(* IEC 61131-3 sources: STAR-PLC-Agent/results/raw/four_group_20261114/star_terra/PUB011/generation/sim_00, 1 file *)

(* ---- test_program.st ---- *)
PROGRAM PLC_PRG
VAR
 BenchStep : UDINT := 0;
 BenchCalls : UDINT := 0;
 BenchDone : BOOL := FALSE;
 BenchUut0 : FB_Task;
 BenchUut1 : FB_Task;
 TraceIn_Mode : ARRAY[0..15] OF BOOL;
 TraceIn_ForwardButton : ARRAY[0..15] OF BOOL;
 TraceIn_ReverseButton : ARRAY[0..15] OF BOOL;
 TraceIn_SensorA : ARRAY[0..15] OF BOOL;
 TraceIn_SensorB : ARRAY[0..15] OF BOOL;
 TraceIn_SensorC : ARRAY[0..15] OF BOOL;
 TraceIn_ButtonA : ARRAY[0..15] OF BOOL;
 TraceIn_ButtonB : ARRAY[0..15] OF BOOL;
 TraceIn_ButtonC : ARRAY[0..15] OF BOOL;
 TraceOut_MotorForward : ARRAY[0..15] OF BOOL;
 TraceOut_MotorReverse : ARRAY[0..15] OF BOOL;
 TraceOut_CompletionLight : ARRAY[0..15] OF BOOL;
END_VAR

IF NOT BenchDone THEN
 CASE BenchStep OF
 0:
   BenchUut0.Mode := TRUE;
   BenchUut0.ForwardButton := FALSE;
   BenchUut0.ReverseButton := FALSE;
   BenchUut0.SensorA := TRUE;
   BenchUut0.SensorB := FALSE;
   BenchUut0.SensorC := FALSE;
   BenchUut0.ButtonA := FALSE;
   BenchUut0.ButtonB := FALSE;
   BenchUut0.ButtonC := FALSE;
   TraceIn_Mode[0] := BenchUut0.Mode;
   TraceIn_ForwardButton[0] := BenchUut0.ForwardButton;
   TraceIn_ReverseButton[0] := BenchUut0.ReverseButton;
   TraceIn_SensorA[0] := BenchUut0.SensorA;
   TraceIn_SensorB[0] := BenchUut0.SensorB;
   TraceIn_SensorC[0] := BenchUut0.SensorC;
   TraceIn_ButtonA[0] := BenchUut0.ButtonA;
   TraceIn_ButtonB[0] := BenchUut0.ButtonB;
   TraceIn_ButtonC[0] := BenchUut0.ButtonC;
   BenchUut0();
   TraceOut_MotorForward[0] := BenchUut0.MotorForward;
   TraceOut_MotorReverse[0] := BenchUut0.MotorReverse;
   TraceOut_CompletionLight[0] := BenchUut0.CompletionLight;
   BenchCalls := BenchCalls + 1;
 1:
   BenchUut0.Mode := TRUE;
   BenchUut0.ForwardButton := FALSE;
   BenchUut0.ReverseButton := FALSE;
   BenchUut0.SensorA := TRUE;
   BenchUut0.SensorB := FALSE;
   BenchUut0.SensorC := FALSE;
   BenchUut0.ButtonA := TRUE;
   BenchUut0.ButtonB := FALSE;
   BenchUut0.ButtonC := FALSE;
   TraceIn_Mode[1] := BenchUut0.Mode;
   TraceIn_ForwardButton[1] := BenchUut0.ForwardButton;
   TraceIn_ReverseButton[1] := BenchUut0.ReverseButton;
   TraceIn_SensorA[1] := BenchUut0.SensorA;
   TraceIn_SensorB[1] := BenchUut0.SensorB;
   TraceIn_SensorC[1] := BenchUut0.SensorC;
   TraceIn_ButtonA[1] := BenchUut0.ButtonA;
   TraceIn_ButtonB[1] := BenchUut0.ButtonB;
   TraceIn_ButtonC[1] := BenchUut0.ButtonC;
   BenchUut0();
   TraceOut_MotorForward[1] := BenchUut0.MotorForward;
   TraceOut_MotorReverse[1] := BenchUut0.MotorReverse;
   TraceOut_CompletionLight[1] := BenchUut0.CompletionLight;
   BenchCalls := BenchCalls + 1;
 2:
   BenchUut0.Mode := TRUE;
   BenchUut0.ForwardButton := FALSE;
   BenchUut0.ReverseButton := FALSE;
   BenchUut0.SensorA := FALSE;
   BenchUut0.SensorB := TRUE;
   BenchUut0.SensorC := FALSE;
   BenchUut0.ButtonA := FALSE;
   BenchUut0.ButtonB := TRUE;
   BenchUut0.ButtonC := FALSE;
   TraceIn_Mode[2] := BenchUut0.Mode;
   TraceIn_ForwardButton[2] := BenchUut0.ForwardButton;
   TraceIn_ReverseButton[2] := BenchUut0.ReverseButton;
   TraceIn_SensorA[2] := BenchUut0.SensorA;
   TraceIn_SensorB[2] := BenchUut0.SensorB;
   TraceIn_SensorC[2] := BenchUut0.SensorC;
   TraceIn_ButtonA[2] := BenchUut0.ButtonA;
   TraceIn_ButtonB[2] := BenchUut0.ButtonB;
   TraceIn_ButtonC[2] := BenchUut0.ButtonC;
   BenchUut0();
   TraceOut_MotorForward[2] := BenchUut0.MotorForward;
   TraceOut_MotorReverse[2] := BenchUut0.MotorReverse;
   TraceOut_CompletionLight[2] := BenchUut0.CompletionLight;
   BenchCalls := BenchCalls + 1;
 3:
   BenchUut0.Mode := TRUE;
   BenchUut0.ForwardButton := FALSE;
   BenchUut0.ReverseButton := FALSE;
   BenchUut0.SensorA := FALSE;
   BenchUut0.SensorB := TRUE;
   BenchUut0.SensorC := FALSE;
   BenchUut0.ButtonA := FALSE;
   BenchUut0.ButtonB := TRUE;
   BenchUut0.ButtonC := FALSE;
   TraceIn_Mode[3] := BenchUut0.Mode;
   TraceIn_ForwardButton[3] := BenchUut0.ForwardButton;
   TraceIn_ReverseButton[3] := BenchUut0.ReverseButton;
   TraceIn_SensorA[3] := BenchUut0.SensorA;
   TraceIn_SensorB[3] := BenchUut0.SensorB;
   TraceIn_SensorC[3] := BenchUut0.SensorC;
   TraceIn_ButtonA[3] := BenchUut0.ButtonA;
   TraceIn_ButtonB[3] := BenchUut0.ButtonB;
   TraceIn_ButtonC[3] := BenchUut0.ButtonC;
   BenchUut0();
   TraceOut_MotorForward[3] := BenchUut0.MotorForward;
   TraceOut_MotorReverse[3] := BenchUut0.MotorReverse;
   TraceOut_CompletionLight[3] := BenchUut0.CompletionLight;
   BenchCalls := BenchCalls + 1;
 4:
   BenchUut0.Mode := TRUE;
   BenchUut0.ForwardButton := FALSE;
   BenchUut0.ReverseButton := FALSE;
   BenchUut0.SensorA := FALSE;
   BenchUut0.SensorB := FALSE;
   BenchUut0.SensorC := TRUE;
   BenchUut0.ButtonA := FALSE;
   BenchUut0.ButtonB := FALSE;
   BenchUut0.ButtonC := TRUE;
   TraceIn_Mode[4] := BenchUut0.Mode;
   TraceIn_ForwardButton[4] := BenchUut0.ForwardButton;
   TraceIn_ReverseButton[4] := BenchUut0.ReverseButton;
   TraceIn_SensorA[4] := BenchUut0.SensorA;
   TraceIn_SensorB[4] := BenchUut0.SensorB;
   TraceIn_SensorC[4] := BenchUut0.SensorC;
   TraceIn_ButtonA[4] := BenchUut0.ButtonA;
   TraceIn_ButtonB[4] := BenchUut0.ButtonB;
   TraceIn_ButtonC[4] := BenchUut0.ButtonC;
   BenchUut0();
   TraceOut_MotorForward[4] := BenchUut0.MotorForward;
   TraceOut_MotorReverse[4] := BenchUut0.MotorReverse;
   TraceOut_CompletionLight[4] := BenchUut0.CompletionLight;
   BenchCalls := BenchCalls + 1;
 5:
   BenchUut0.Mode := TRUE;
   BenchUut0.ForwardButton := FALSE;
   BenchUut0.ReverseButton := FALSE;
   BenchUut0.SensorA := FALSE;
   BenchUut0.SensorB := FALSE;
   BenchUut0.SensorC := TRUE;
   BenchUut0.ButtonA := FALSE;
   BenchUut0.ButtonB := FALSE;
   BenchUut0.ButtonC := TRUE;
   TraceIn_Mode[5] := BenchUut0.Mode;
   TraceIn_ForwardButton[5] := BenchUut0.ForwardButton;
   TraceIn_ReverseButton[5] := BenchUut0.ReverseButton;
   TraceIn_SensorA[5] := BenchUut0.SensorA;
   TraceIn_SensorB[5] := BenchUut0.SensorB;
   TraceIn_SensorC[5] := BenchUut0.SensorC;
   TraceIn_ButtonA[5] := BenchUut0.ButtonA;
   TraceIn_ButtonB[5] := BenchUut0.ButtonB;
   TraceIn_ButtonC[5] := BenchUut0.ButtonC;
   BenchUut0();
   TraceOut_MotorForward[5] := BenchUut0.MotorForward;
   TraceOut_MotorReverse[5] := BenchUut0.MotorReverse;
   TraceOut_CompletionLight[5] := BenchUut0.CompletionLight;
   BenchCalls := BenchCalls + 1;
 6:
   BenchUut0.Mode := TRUE;
   BenchUut0.ForwardButton := FALSE;
   BenchUut0.ReverseButton := FALSE;
   BenchUut0.SensorA := FALSE;
   BenchUut0.SensorB := FALSE;
   BenchUut0.SensorC := TRUE;
   BenchUut0.ButtonA := FALSE;
   BenchUut0.ButtonB := FALSE;
   BenchUut0.ButtonC := FALSE;
   TraceIn_Mode[6] := BenchUut0.Mode;
   TraceIn_ForwardButton[6] := BenchUut0.ForwardButton;
   TraceIn_ReverseButton[6] := BenchUut0.ReverseButton;
   TraceIn_SensorA[6] := BenchUut0.SensorA;
   TraceIn_SensorB[6] := BenchUut0.SensorB;
   TraceIn_SensorC[6] := BenchUut0.SensorC;
   TraceIn_ButtonA[6] := BenchUut0.ButtonA;
   TraceIn_ButtonB[6] := BenchUut0.ButtonB;
   TraceIn_ButtonC[6] := BenchUut0.ButtonC;
   BenchUut0();
   TraceOut_MotorForward[6] := BenchUut0.MotorForward;
   TraceOut_MotorReverse[6] := BenchUut0.MotorReverse;
   TraceOut_CompletionLight[6] := BenchUut0.CompletionLight;
   BenchCalls := BenchCalls + 1;
 7:
   BenchUut0.Mode := TRUE;
   BenchUut0.ForwardButton := FALSE;
   BenchUut0.ReverseButton := FALSE;
   BenchUut0.SensorA := FALSE;
   BenchUut0.SensorB := FALSE;
   BenchUut0.SensorC := FALSE;
   BenchUut0.ButtonA := FALSE;
   BenchUut0.ButtonB := FALSE;
   BenchUut0.ButtonC := FALSE;
   TraceIn_Mode[7] := BenchUut0.Mode;
   TraceIn_ForwardButton[7] := BenchUut0.ForwardButton;
   TraceIn_ReverseButton[7] := BenchUut0.ReverseButton;
   TraceIn_SensorA[7] := BenchUut0.SensorA;
   TraceIn_SensorB[7] := BenchUut0.SensorB;
   TraceIn_SensorC[7] := BenchUut0.SensorC;
   TraceIn_ButtonA[7] := BenchUut0.ButtonA;
   TraceIn_ButtonB[7] := BenchUut0.ButtonB;
   TraceIn_ButtonC[7] := BenchUut0.ButtonC;
   BenchUut0();
   TraceOut_MotorForward[7] := BenchUut0.MotorForward;
   TraceOut_MotorReverse[7] := BenchUut0.MotorReverse;
   TraceOut_CompletionLight[7] := BenchUut0.CompletionLight;
   BenchCalls := BenchCalls + 1;
 8:
   BenchUut1.Mode := FALSE;
   BenchUut1.ForwardButton := TRUE;
   BenchUut1.ReverseButton := FALSE;
   BenchUut1.SensorA := FALSE;
   BenchUut1.SensorB := FALSE;
   BenchUut1.SensorC := FALSE;
   BenchUut1.ButtonA := FALSE;
   BenchUut1.ButtonB := FALSE;
   BenchUut1.ButtonC := FALSE;
   TraceIn_Mode[8] := BenchUut1.Mode;
   TraceIn_ForwardButton[8] := BenchUut1.ForwardButton;
   TraceIn_ReverseButton[8] := BenchUut1.ReverseButton;
   TraceIn_SensorA[8] := BenchUut1.SensorA;
   TraceIn_SensorB[8] := BenchUut1.SensorB;
   TraceIn_SensorC[8] := BenchUut1.SensorC;
   TraceIn_ButtonA[8] := BenchUut1.ButtonA;
   TraceIn_ButtonB[8] := BenchUut1.ButtonB;
   TraceIn_ButtonC[8] := BenchUut1.ButtonC;
   BenchUut1();
   TraceOut_MotorForward[8] := BenchUut1.MotorForward;
   TraceOut_MotorReverse[8] := BenchUut1.MotorReverse;
   TraceOut_CompletionLight[8] := BenchUut1.CompletionLight;
   BenchCalls := BenchCalls + 1;
 9:
   BenchUut1.Mode := FALSE;
   BenchUut1.ForwardButton := TRUE;
   BenchUut1.ReverseButton := TRUE;
   BenchUut1.SensorA := FALSE;
   BenchUut1.SensorB := FALSE;
   BenchUut1.SensorC := FALSE;
   BenchUut1.ButtonA := FALSE;
   BenchUut1.ButtonB := FALSE;
   BenchUut1.ButtonC := FALSE;
   TraceIn_Mode[9] := BenchUut1.Mode;
   TraceIn_ForwardButton[9] := BenchUut1.ForwardButton;
   TraceIn_ReverseButton[9] := BenchUut1.ReverseButton;
   TraceIn_SensorA[9] := BenchUut1.SensorA;
   TraceIn_SensorB[9] := BenchUut1.SensorB;
   TraceIn_SensorC[9] := BenchUut1.SensorC;
   TraceIn_ButtonA[9] := BenchUut1.ButtonA;
   TraceIn_ButtonB[9] := BenchUut1.ButtonB;
   TraceIn_ButtonC[9] := BenchUut1.ButtonC;
   BenchUut1();
   TraceOut_MotorForward[9] := BenchUut1.MotorForward;
   TraceOut_MotorReverse[9] := BenchUut1.MotorReverse;
   TraceOut_CompletionLight[9] := BenchUut1.CompletionLight;
   BenchCalls := BenchCalls + 1;
 10:
   BenchUut1.Mode := FALSE;
   BenchUut1.ForwardButton := FALSE;
   BenchUut1.ReverseButton := TRUE;
   BenchUut1.SensorA := FALSE;
   BenchUut1.SensorB := FALSE;
   BenchUut1.SensorC := FALSE;
   BenchUut1.ButtonA := FALSE;
   BenchUut1.ButtonB := FALSE;
   BenchUut1.ButtonC := FALSE;
   TraceIn_Mode[10] := BenchUut1.Mode;
   TraceIn_ForwardButton[10] := BenchUut1.ForwardButton;
   TraceIn_ReverseButton[10] := BenchUut1.ReverseButton;
   TraceIn_SensorA[10] := BenchUut1.SensorA;
   TraceIn_SensorB[10] := BenchUut1.SensorB;
   TraceIn_SensorC[10] := BenchUut1.SensorC;
   TraceIn_ButtonA[10] := BenchUut1.ButtonA;
   TraceIn_ButtonB[10] := BenchUut1.ButtonB;
   TraceIn_ButtonC[10] := BenchUut1.ButtonC;
   BenchUut1();
   TraceOut_MotorForward[10] := BenchUut1.MotorForward;
   TraceOut_MotorReverse[10] := BenchUut1.MotorReverse;
   TraceOut_CompletionLight[10] := BenchUut1.CompletionLight;
   BenchCalls := BenchCalls + 1;
 11:
   BenchUut1.Mode := TRUE;
   BenchUut1.ForwardButton := FALSE;
   BenchUut1.ReverseButton := TRUE;
   BenchUut1.SensorA := TRUE;
   BenchUut1.SensorB := FALSE;
   BenchUut1.SensorC := FALSE;
   BenchUut1.ButtonA := TRUE;
   BenchUut1.ButtonB := FALSE;
   BenchUut1.ButtonC := FALSE;
   TraceIn_Mode[11] := BenchUut1.Mode;
   TraceIn_ForwardButton[11] := BenchUut1.ForwardButton;
   TraceIn_ReverseButton[11] := BenchUut1.ReverseButton;
   TraceIn_SensorA[11] := BenchUut1.SensorA;
   TraceIn_SensorB[11] := BenchUut1.SensorB;
   TraceIn_SensorC[11] := BenchUut1.SensorC;
   TraceIn_ButtonA[11] := BenchUut1.ButtonA;
   TraceIn_ButtonB[11] := BenchUut1.ButtonB;
   TraceIn_ButtonC[11] := BenchUut1.ButtonC;
   BenchUut1();
   TraceOut_MotorForward[11] := BenchUut1.MotorForward;
   TraceOut_MotorReverse[11] := BenchUut1.MotorReverse;
   TraceOut_CompletionLight[11] := BenchUut1.CompletionLight;
   BenchCalls := BenchCalls + 1;
 12:
   BenchUut1.Mode := TRUE;
   BenchUut1.ForwardButton := FALSE;
   BenchUut1.ReverseButton := TRUE;
   BenchUut1.SensorA := FALSE;
   BenchUut1.SensorB := FALSE;
   BenchUut1.SensorC := FALSE;
   BenchUut1.ButtonA := FALSE;
   BenchUut1.ButtonB := FALSE;
   BenchUut1.ButtonC := FALSE;
   TraceIn_Mode[12] := BenchUut1.Mode;
   TraceIn_ForwardButton[12] := BenchUut1.ForwardButton;
   TraceIn_ReverseButton[12] := BenchUut1.ReverseButton;
   TraceIn_SensorA[12] := BenchUut1.SensorA;
   TraceIn_SensorB[12] := BenchUut1.SensorB;
   TraceIn_SensorC[12] := BenchUut1.SensorC;
   TraceIn_ButtonA[12] := BenchUut1.ButtonA;
   TraceIn_ButtonB[12] := BenchUut1.ButtonB;
   TraceIn_ButtonC[12] := BenchUut1.ButtonC;
   BenchUut1();
   TraceOut_MotorForward[12] := BenchUut1.MotorForward;
   TraceOut_MotorReverse[12] := BenchUut1.MotorReverse;
   TraceOut_CompletionLight[12] := BenchUut1.CompletionLight;
   BenchCalls := BenchCalls + 1;
 13:
   BenchUut1.Mode := FALSE;
   BenchUut1.ForwardButton := FALSE;
   BenchUut1.ReverseButton := TRUE;
   BenchUut1.SensorA := FALSE;
   BenchUut1.SensorB := FALSE;
   BenchUut1.SensorC := FALSE;
   BenchUut1.ButtonA := FALSE;
   BenchUut1.ButtonB := FALSE;
   BenchUut1.ButtonC := FALSE;
   TraceIn_Mode[13] := BenchUut1.Mode;
   TraceIn_ForwardButton[13] := BenchUut1.ForwardButton;
   TraceIn_ReverseButton[13] := BenchUut1.ReverseButton;
   TraceIn_SensorA[13] := BenchUut1.SensorA;
   TraceIn_SensorB[13] := BenchUut1.SensorB;
   TraceIn_SensorC[13] := BenchUut1.SensorC;
   TraceIn_ButtonA[13] := BenchUut1.ButtonA;
   TraceIn_ButtonB[13] := BenchUut1.ButtonB;
   TraceIn_ButtonC[13] := BenchUut1.ButtonC;
   BenchUut1();
   TraceOut_MotorForward[13] := BenchUut1.MotorForward;
   TraceOut_MotorReverse[13] := BenchUut1.MotorReverse;
   TraceOut_CompletionLight[13] := BenchUut1.CompletionLight;
   BenchCalls := BenchCalls + 1;
 14:
   BenchUut1.Mode := TRUE;
   BenchUut1.ForwardButton := FALSE;
   BenchUut1.ReverseButton := FALSE;
   BenchUut1.SensorA := FALSE;
   BenchUut1.SensorB := TRUE;
   BenchUut1.SensorC := FALSE;
   BenchUut1.ButtonA := FALSE;
   BenchUut1.ButtonB := TRUE;
   BenchUut1.ButtonC := FALSE;
   TraceIn_Mode[14] := BenchUut1.Mode;
   TraceIn_ForwardButton[14] := BenchUut1.ForwardButton;
   TraceIn_ReverseButton[14] := BenchUut1.ReverseButton;
   TraceIn_SensorA[14] := BenchUut1.SensorA;
   TraceIn_SensorB[14] := BenchUut1.SensorB;
   TraceIn_SensorC[14] := BenchUut1.SensorC;
   TraceIn_ButtonA[14] := BenchUut1.ButtonA;
   TraceIn_ButtonB[14] := BenchUut1.ButtonB;
   TraceIn_ButtonC[14] := BenchUut1.ButtonC;
   BenchUut1();
   TraceOut_MotorForward[14] := BenchUut1.MotorForward;
   TraceOut_MotorReverse[14] := BenchUut1.MotorReverse;
   TraceOut_CompletionLight[14] := BenchUut1.CompletionLight;
   BenchCalls := BenchCalls + 1;
 15:
   BenchUut1.Mode := TRUE;
   BenchUut1.ForwardButton := FALSE;
   BenchUut1.ReverseButton := FALSE;
   BenchUut1.SensorA := TRUE;
   BenchUut1.SensorB := FALSE;
   BenchUut1.SensorC := FALSE;
   BenchUut1.ButtonA := TRUE;
   BenchUut1.ButtonB := FALSE;
   BenchUut1.ButtonC := FALSE;
   TraceIn_Mode[15] := BenchUut1.Mode;
   TraceIn_ForwardButton[15] := BenchUut1.ForwardButton;
   TraceIn_ReverseButton[15] := BenchUut1.ReverseButton;
   TraceIn_SensorA[15] := BenchUut1.SensorA;
   TraceIn_SensorB[15] := BenchUut1.SensorB;
   TraceIn_SensorC[15] := BenchUut1.SensorC;
   TraceIn_ButtonA[15] := BenchUut1.ButtonA;
   TraceIn_ButtonB[15] := BenchUut1.ButtonB;
   TraceIn_ButtonC[15] := BenchUut1.ButtonC;
   BenchUut1();
   TraceOut_MotorForward[15] := BenchUut1.MotorForward;
   TraceOut_MotorReverse[15] := BenchUut1.MotorReverse;
   TraceOut_CompletionLight[15] := BenchUut1.CompletionLight;
   BenchCalls := BenchCalls + 1;
 END_CASE;
 BenchStep := BenchStep + 1;
 IF BenchStep >= 16 THEN BenchDone := TRUE; END_IF;
END_IF;
END_PROGRAM
